Fanuc KAREL source: kb00073.compact.KL

PROGRAM KB00073
%STACKSIZE=65535
%PRIORITY=65535
%NOLOCKGROUP
VAR
P1 : INTEGER
P2 : STRING[80]
BEGIN
P1=1
P2='A'
FORCE_LINK(P1,P2)
END KB00073
